Staubli VAL3: HMI_TRAJ.dtx

mdesc mNomSpeed
string sUsingLib
string sList
bool bBack
bool bBool[12]
string sPageIndex
string sPageNum
num nPageIndex
num nPageNum
string sNewName
string sFrameList
string sToolList
bool bConfirm
bool bCancel
num nMoveID
string sSelFrame
string sSelTool
string sSelTraj
bool bRefresh
bool bToSave
public trajItem tEditItem
  [0]
    num nFrameIndex
    num nToolIndex
    string sID
    num nMoveID
    pointItem pPointItem
      [0]
        pointRx pPointRx[2]
        jointRx jJointRx
        paraItem pParaItem
          [0]
            mdesc mMdesc
            num nMoveType
            num nActionIndex
            num nPercentage
            ifItem iIfItem
              [0]
                num nSigType[3]
                num nSigIndex[3]
                num nValue[3]
                bool bANDOR[2]
            num nDelay
            num nSigValue
            bool bSafePoint
        string sID
        bool bMarked
        pointRx pInter
string sTrajList
string sTrajList1
string sSessionList
num nIDIsExit
